(* IEC 61131-3 sources: kns-pump-station/tests/POUs/Log/FB_EventLogCsv_Test, 14 files *)

(* ---- FB_EventLogCsv_Test.decl.st ---- *)
// Назначение: набор coUnit для FB_EventLogCsv и F_EventCsvLine — формат строки CSV; выгрузка через CAA File в
//             рантайме (многоцикловые тесты): заголовок и все строки снимка, пустой снимок, чтение файла назад
//             и побайтное сравнение (как зонд Z1 архитектуры), ошибка на несуществующем каталоге. Файлы —
//             в рабочем каталоге рантайма (относительные имена kns_test_*.csv).
// Автор:      kr0nsch
// Версия:     0.1.0
// Документ:   docs/DESIGN.md, разделы 9.2, 14.1
FUNCTION_BLOCK FB_EventLogCsv_Test EXTENDS coUnit.FB_TestSuite
VAR CONSTANT
    POLLS_MAX : UINT := 1000;       // предел вызовов теста на выгрузку (≈ 10 с при TestTask 10 мс)
    READ_BUF_LEN : UINT := 4096;    // буфер чтения файла назад
END_VAR

(* ---- AppendExpected.method.decl.st ---- *)
// Дописать ASCII-байты строки в буфер ожидаемого содержимого
METHOD PRIVATE AppendExpected
VAR_INPUT
    sText : STRING(GVL_Const.LOG_CSV_LINE_LEN);
END_VAR
VAR_IN_OUT
    abBuf  : ARRAY[0..READ_BUF_LEN - 1] OF BYTE;
    udiLen : UDINT;
END_VAR
VAR
    pChar : POINTER TO BYTE;        // очередной символ строки
    iI    : INT;                    // номер символа
END_VAR

(* ---- AppendExpected.method.impl.st ---- *)
pChar := ADR(sText);
FOR iI := 1 TO LEN(sText) DO
    IF udiLen < READ_BUF_LEN THEN
        abBuf[udiLen] := pChar^;
        udiLen := udiLen + 1;
    END_IF
    pChar := pChar + 1;
END_FOR

(* ---- EmptySnapshotHeaderOnly.method.decl.st ---- *)
// Пустой снимок: файл с одним заголовком, Done, строк 0
METHOD PRIVATE EmptySnapshotHeaderOnly
VAR_INST
    fbLog    : FB_EventLog;         // пустой журнал
    fbCsv    : FB_EventLogCsv;      // проверяемая выгрузка
    uiPolls : UINT;                // вызовов теста с начала
END_VAR

(* ---- EmptySnapshotHeaderOnly.method.impl.st ---- *)
coUnit.TEST('EventLogCsv_EmptySnapshotHeaderOnly');

IF uiPolls = 0 THEN
    fbLog.TakeSnapshot();
END_IF
fbCsv(xExecute := TRUE, sFileName := 'kns_test_events_empty.csv', fbLog := fbLog);
uiPolls := uiPolls + 1;
IF fbCsv.xDone OR fbCsv.xError OR uiPolls >= POLLS_MAX THEN
    AssertTrue(Condition := fbCsv.xDone AND NOT fbCsv.xError, Message := 'header-only export done');
    AssertEquals_UINT(Expected := 0, Actual := fbCsv.uiLines, Message := 'no data lines');
    coUnit.TEST_FINISHED();
END_IF

(* ---- ErrorOnBadPathReported.method.decl.st ---- *)
// Пустое имя файла: открытие не удаётся — Error, код FILE.ERROR не 0, строк 0 (несуществующий каталог
// CAA File на Control Win создаёт сам — проверено прогоном)
METHOD PRIVATE ErrorOnBadPathReported
VAR_INST
    fbLog    : FB_EventLog;         // журнал со снимком
    fbCsv    : FB_EventLogCsv;      // проверяемая выгрузка
    uiPolls : UINT;                // вызовов теста с начала
END_VAR

(* ---- ErrorOnBadPathReported.method.impl.st ---- *)
coUnit.TEST('EventLogCsv_ErrorOnBadPathReported');

IF uiPolls = 0 THEN
    fbLog.LogEvent(eEvent := E_StationEvent.PlcStart, rValue := 0.0);
    fbLog.TakeSnapshot();
END_IF
fbCsv(xExecute := TRUE, sFileName := '', fbLog := fbLog);
uiPolls := uiPolls + 1;
IF fbCsv.xDone OR fbCsv.xError OR uiPolls >= POLLS_MAX THEN
    AssertTrue(Condition := fbCsv.xError, Message := 'error reported');
    AssertFalse(Condition := fbCsv.xDone, Message := 'not done');
    AssertTrue(Condition := fbCsv.eState = E_LogExportState.Error, Message := 'state Error');
    AssertTrue(Condition := fbCsv.udiError <> 0, Message := 'CAA File error code');
    AssertEquals_UINT(Expected := 0, Actual := fbCsv.uiLines, Message := 'no lines');
    coUnit.TEST_FINISHED();
END_IF

(* ---- EventCsvLineFormat.method.decl.st ---- *)
// Строка CSV: тревога (UTC, код P101.FTS, числа перечислений) и событие станции без часов (пустое время);
// значение — REAL_TO_STRING (3.0 → «3.0», проверено прогоном)
METHOD PRIVATE EventCsvLineFormat
VAR
    stRec : ST_EventRecord;         // запись журнала
END_VAR

(* ---- ReadBackMatchesSnapshot.method.decl.st ---- *)
// Выгрузка 12 записей, затем файл читается назад (FILE.Open MREAD, Read, Close): длина и байты совпадают с
// заголовком и строками F_EventCsvLine снимка
METHOD PRIVATE ReadBackMatchesSnapshot
VAR_INST
    fbLog     : FB_EventLog;        // журнал со снимком
    fbCsv     : FB_EventLogCsv;     // проверяемая выгрузка
    fbOpen    : FILE.Open;          // чтение назад
    fbRead    : FILE.Read;
    fbClose   : FILE.Close;
    abRead    : ARRAY[0..READ_BUF_LEN - 1] OF BYTE;   // прочитанный файл
    abExp     : ARRAY[0..READ_BUF_LEN - 1] OF BYTE;   // ожидаемое содержимое
    udiExpLen : UDINT;              // байт ожидаемого содержимого
    udiReadLen : UDINT;             // байт прочитано
    uiPolls  : UINT;               // вызовов теста с начала
    iStep     : INT;                // 0 — запись, 1 — открыть, 2 — читать, 3 — закрыть, 4 — сравнить
    xReadError : BOOL;              // ошибка CAA File при чтении назад
END_VAR
VAR
    fbTime  : PL.FB_FakeTime;       // подменное время
    stRec   : ST_EventRecord;       // запись снимка
    uiI     : UINT;                 // номер записи
    udiDiff : UDINT;                // байт, отличных от ожидаемых
    udiK    : UDINT;                // номер байта
END_VAR

(* ---- ReadBackMatchesSnapshot.method.impl.st ---- *)
coUnit.TEST('EventLogCsv_ReadBackMatchesSnapshot');

IF uiPolls = 0 THEN
    fbLog.itfTime := fbTime;
    FOR uiI := 1 TO 12 DO
        fbTime.Advance(tStep := T#1S);
        fbLog.LogEvent(eEvent := E_StationEvent.LeadChanged, rValue := UINT_TO_REAL(uiI));
    END_FOR
    fbLog.TakeSnapshot();
    // ожидаемое содержимое: заголовок и строки снимка
    AppendExpected(sText := GVL_Const.LOG_CSV_HEADER, abBuf := abExp, udiLen := udiExpLen);
    FOR uiI := 1 TO fbLog.SnapshotCount DO
        fbLog.GetSnapshotRecord(uiIndex := uiI - 1, stRecord => stRec);
        AppendExpected(sText := F_EventCsvLine(stRecord := stRec), abBuf := abExp, udiLen := udiExpLen);
    END_FOR
END_IF
uiPolls := uiPolls + 1;
CASE iStep OF
    0:
        fbCsv(xExecute := TRUE, sFileName := 'kns_test_events_read.csv', fbLog := fbLog);
        IF fbCsv.xDone OR fbCsv.xError THEN
            iStep := 1;
        END_IF
    1:
        fbOpen(xExecute := TRUE, sFileName := 'kns_test_events_read.csv', eFileMode := FILE.MODE.MREAD,
               xExclusive := FALSE);
        IF fbOpen.xDone THEN
            iStep := 2;
        ELSIF fbOpen.xError THEN
            xReadError := TRUE;
            iStep := 4;
        END_IF
    2:
        fbRead(xExecute := TRUE, hFile := fbOpen.hFile, pBuffer := ADR(abRead), szBuffer := SIZEOF(abRead),
               udiTimeOut := GVL_Const.LOG_CSV_TIMEOUT_US);
        IF fbRead.xDone OR fbRead.xError THEN
            xReadError := fbRead.xError;
            udiReadLen := TO_UDINT(fbRead.szSize);
            iStep := 3;
        END_IF
    3:
        fbClose(xExecute := TRUE, hFile := fbOpen.hFile);
        IF fbClose.xDone OR fbClose.xError THEN
            iStep := 4;
        END_IF
END_CASE
IF iStep = 4 OR uiPolls >= POLLS_MAX THEN
    AssertTrue(Condition := fbCsv.xDone, Message := 'export done');
    AssertFalse(Condition := xReadError, Message := 'file read back without CAA File error');
    AssertEquals_UDINT(Expected := udiExpLen, Actual := udiReadLen, Message := 'file length = expected');
    udiDiff := 0;
    FOR udiK := 1 TO MIN(udiExpLen, udiReadLen) DO
        IF abRead[udiK - 1] <> abExp[udiK - 1] THEN
            udiDiff := udiDiff + 1;
        END_IF
    END_FOR
    AssertEquals_UDINT(Expected := 0, Actual := udiDiff, Message := 'file bytes = header + snapshot lines');
    AssertTrue(Condition := udiExpLen > 0, Message := 'expected content not empty');
    coUnit.TEST_FINISHED();
END_IF

(* ---- SlowTaskRequestHandshake.method.decl.st ---- *)
// Обмен MainTask ↔ SlowTask через PRG_Slow и GVL_Log: запрос снимается, как только выгрузка началась
// (Writing); итог — Done и число строк; запрос сразу после Done (до следующего цикла SlowTask) запускает
// вторую выгрузку, а не теряется
METHOD PRIVATE SlowTaskRequestHandshake
VAR_INST
    fbTime  : PL.FB_FakeTime;       // время журнала (переживает циклы теста)
    uiPolls : UINT;                 // вызовов теста с начала
    iStep   : INT;                  // 0 — первый запрос, 1 — первая выгрузка, 2 — вторая выгрузка, 3 — итог
    xSecond : BOOL;                 // вторая выгрузка началась (Writing)
END_VAR
VAR
    uiI : UINT;                     // номер события
END_VAR

(* ---- SlowTaskRequestHandshake.method.impl.st ---- *)
coUnit.TEST('EventLogCsv_SlowTaskRequestHandshake');

uiPolls := uiPolls + 1;
CASE iStep OF
    0:
        GVL_Log.fbEventLog.itfTime := fbTime;
        FOR uiI := 1 TO 3 DO
            GVL_Log.fbEventLog.LogEvent(eEvent := E_StationEvent.CfgChanged, rValue := UINT_TO_REAL(uiI));
        END_FOR
        GVL_Log.fbEventLog.TakeSnapshot();
        GVL_Log.xExportReq := TRUE;
        PRG_Slow();
        AssertTrue(Condition := GVL_Log.eExportState = E_LogExportState.Writing, Message := 'first export started');
        AssertFalse(Condition := GVL_Log.xExportReq, Message := 'request taken when export starts');
        iStep := 1;
    1:
        PRG_Slow();
        IF GVL_Log.eExportState = E_LogExportState.Done OR GVL_Log.eExportState = E_LogExportState.Error THEN
            AssertTrue(Condition := GVL_Log.eExportState = E_LogExportState.Done, Message := 'first export done');
            AssertEquals_UINT(Expected := 3, Actual := GVL_Log.uiExportLines, Message := 'first export: 3 lines');
            // MainTask видит Done и сразу ставит новый запрос — до следующего цикла SlowTask
            GVL_Log.fbEventLog.LogEvent(eEvent := E_StationEvent.CfgChanged, rValue := 4.0);
            GVL_Log.fbEventLog.LogEvent(eEvent := E_StationEvent.CfgChanged, rValue := 5.0);
            GVL_Log.fbEventLog.TakeSnapshot();
            GVL_Log.xExportReq := TRUE;
            PRG_Slow();
            xSecond := GVL_Log.eExportState = E_LogExportState.Writing;
            AssertTrue(Condition := xSecond, Message := 'request right after Done starts second export');
            AssertFalse(Condition := GVL_Log.xExportReq, Message := 'second request taken');
            iStep := SEL(xSecond, 3, 2);
        END_IF
    2:
        PRG_Slow();
        IF GVL_Log.eExportState = E_LogExportState.Done OR GVL_Log.eExportState = E_LogExportState.Error THEN
            AssertTrue(Condition := GVL_Log.eExportState = E_LogExportState.Done, Message := 'second export done');
            AssertEquals_UINT(Expected := 5, Actual := GVL_Log.uiExportLines, Message := 'second export: 5 lines');
            AssertFalse(Condition := GVL_Log.xExportReq, Message := 'no request left');
            iStep := 3;
        END_IF
END_CASE
IF iStep = 3 OR uiPolls >= POLLS_MAX THEN
    AssertTrue(Condition := iStep = 3, Message := 'handshake finished in time');
    GVL_Log.fbEventLog.itfTime := 0;
    coUnit.TEST_FINISHED();
END_IF

(* ---- WritesHeaderAndAllLines.method.decl.st ---- *)
// 25 записей (три порции FILE.Write по 10 строк): выгрузка завершается Done, строк 25, ошибки нет
METHOD PRIVATE WritesHeaderAndAllLines
VAR_INST
    fbLog    : FB_EventLog;         // журнал со снимком
    fbCsv    : FB_EventLogCsv;      // проверяемая выгрузка
    uiPolls : UINT;                // вызовов теста с начала
    xStarted : BOOL;                // записи и снимок готовы
END_VAR
VAR
    fbTime : PL.FB_FakeTime;        // подменное время
    uiI    : UINT;                  // номер события
END_VAR

(* ---- WritesHeaderAndAllLines.method.impl.st ---- *)
coUnit.TEST('EventLogCsv_WritesHeaderAndAllLines');

IF NOT xStarted THEN
    fbLog.itfTime := fbTime;
    FOR uiI := 1 TO 25 DO
        fbLog.LogEvent(eEvent := E_StationEvent.CfgChanged, rValue := UINT_TO_REAL(uiI));
    END_FOR
    fbLog.TakeSnapshot();
    xStarted := TRUE;
END_IF
fbCsv(xExecute := TRUE, sFileName := 'kns_test_events_all.csv', fbLog := fbLog);
uiPolls := uiPolls + 1;
IF fbCsv.xDone OR fbCsv.xError OR uiPolls >= POLLS_MAX THEN
    AssertTrue(Condition := fbCsv.xDone, Message := 'export done');
    AssertFalse(Condition := fbCsv.xError, Message := 'no error');
    AssertTrue(Condition := fbCsv.eState = E_LogExportState.Done, Message := 'state Done');
    AssertEquals_UINT(Expected := 25, Actual := fbCsv.uiLines, Message := '25 lines');
    AssertEquals_UDINT(Expected := 0, Actual := fbCsv.udiError, Message := 'error code 0');
    coUnit.TEST_FINISHED();
END_IF
